# B&R Automation Studio project lab3
Automation Studio 4.5.2.102; technology packages: Acp10Arnc0 5.2.1

## Configuration Config1

CPU 4PP065.0571-P74, AutomationRuntime D4.52, Build 4.1.2, Vc V4.52.0, Safety 1.6

### Task classes (Cpu.sw)
```
Cyclic#1 (cycle 2000 us, tolerance 0 us):
  SDCAxisCtr <- SDCAxisCtrlX.prg
DataObjects: Acp10sys
NcDataObjects: acp10etxen <- acp10etxen.dob, Axis_Xa <- Axis_Xobj.Axis_Xa.dob, Axis_Xi <- Axis_Xobj.Axis_Xi.dob
Binaries: TCData, udbdef, ashwd, Role, User, sysconf, ashwac, asfw, arconfig, iomap, acp10cfg, Acp10map1, Acp10map
Libraries: Acp10man, Acp10par, NcGlobal, Acp10sdc, Acp10_MC, brsystem, sys_lib, runtime, AsBrStr, Acp10sim, AsIOTime, MotorContr, asstring, astime, fileio, powerlnk, asieccon
```

### Hardware
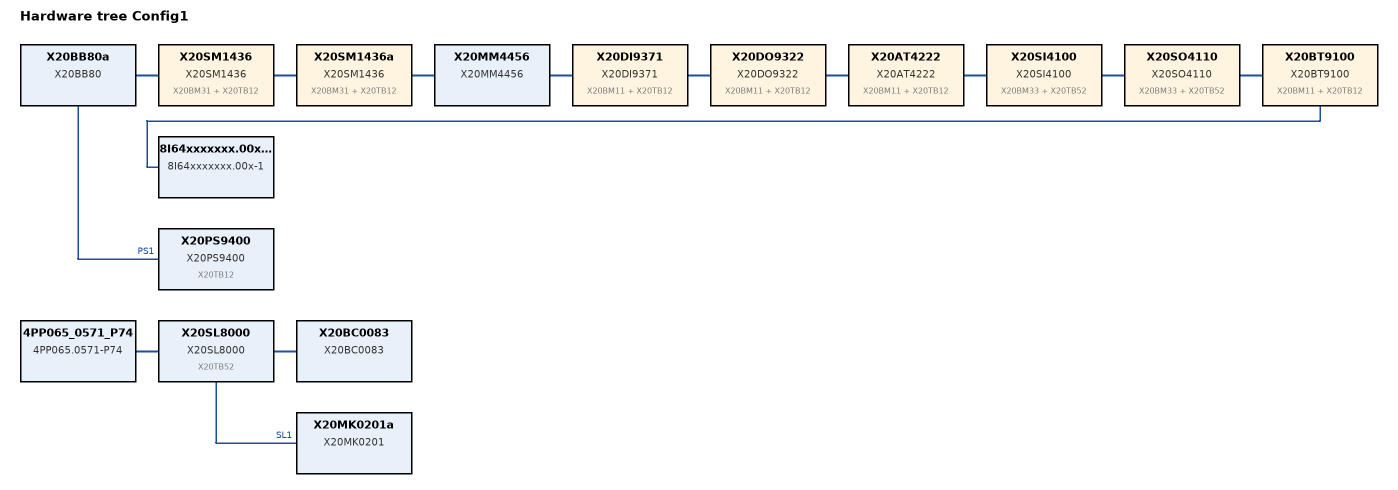
```
4PP065_0571_P74 : 4PP065.0571-P74 v1.1.2.0
  Connector IF5:
    ActivateDevice = 1
    Mode = Manual
    InternetAddress = 10.0.1.10
    SubnetMask = 255.255.255.0
  ConfigurationID = labBR
  TimerDeviceType = EPLX2X
  TimerDevice = 4PP065_0571_P74.IF4
  TaskClassIdleTime = 2000
  Cyclic1Duration = 2000
  Cyclic1Tolerance = 0
  Cyclic1Output = 1
8I64xxxxxxx.00x-1 : 8I64xxxxxxx.00x-1 v2.1.3.0  [X2X1 -> X20BT9100.X2X1 [Cable Type=X2XCable, Length=10, Version=1.0.0.2]]
  packedETAD = packed
  packedETI = packed
  packedCMDD = packed
  ACC = 30
  DEC = 30
  UNS = 220
  NCR = 10
  NSP = 890
  COS = 64
  RSC = 33000
X20AT4222 : X20AT4222 v1.2.3.0  [SS1 -> X20TB12f.SS; SL -> X20BM11c.SL1]
X20BB80a : X20BB80 v1.0.2.0
X20BC0083 : X20BC0083 v2.9.0.0  [PLK1 -> X20SL8000.PLK2 (NodeNumber=2) [Cable Type=PowerlinkCable, Length=10, Version=1.0.0.2]; SL -> X20BB80a.SL1]
X20BM11a : X20BM11 v1.0.0.1  [X2X1 -> X20MM4456.X2X2]
X20BM11b : X20BM11 v1.0.0.1  [X2X1 -> X20BM11a.X2X2]
X20BM11c : X20BM11 v1.0.0.1  [X2X1 -> X20BM11b.X2X2]
X20BM11d : X20BM11 v1.0.0.1  [X2X1 -> X20BM33b.X2X2]
X20BM31a : X20BM31 v1.0.0.1  [X2X1 -> X20BB80a.IF1]
X20BM31b : X20BM31 v1.0.0.1  [X2X1 -> X20BM31a.X2X2]
X20BM33a : X20BM33 v1.0.0.4  [X2X1 -> X20BM11c.X2X2]
X20BM33b : X20BM33 v1.0.0.4  [X2X1 -> X20BM33a.X2X2]
X20BT9100 : X20BT9100 v1.0.3.0  [SS1 -> X20TB12g.SS; SL -> X20BM11d.SL1]
X20DI9371 : X20DI9371 v1.0.2.0  [SS1 -> X20TB12d.SS; SL -> X20BM11a.SL1]
X20DO9322 : X20DO9322 v1.0.3.0  [SS1 -> X20TB12e.SS; SL -> X20BM11b.SL1]
X20MK0201a : X20MK0201 v1.0.0.0  [SL -> X20SL8000.SL1]
X20MM4456 : X20MM4456 v1.1.5.0  [X2X1 -> X20BM31b.X2X2]
X20PS9400 : X20PS9400 v1.8.0.0  [SS1 -> X20TB12b.SS; PS -> X20BB80a.PS1]
X20SI4100 : X20SI4100 v1.10.1.1  [SS1 -> X20TB52b.SS; SL -> X20BM33a.SL1]
X20SL8000 : X20SL8000 v1.6.5.2  [PLK1 -> 4PP065_0571_P74.IF4 (NodeNumber=1) [Cable Type=PowerlinkCable, Length=10, Version=1.0.0.2]; PLK2 -> X20BC0083.PLK1 (NodeNumber=1) [Cable Type=PowerlinkCable, Length=10, Version=1.0.0.2]; SS1 -> X20TB52a.SS]
  SafeProject = SafeLOGIC-1
  SafeDesigner = 3.0.18.3402403
X20SM1436 : X20SM1436 v2.3.0.0  [SS1 -> X20TB12a.SS; SL -> X20BM31a.SL1]
X20SM1436a : X20SM1436 v2.3.0.0  [SS1 -> X20TB12c.SS; SL -> X20BM31b.SL1]
X20SO4110 : X20SO4110 v1.10.1.1  [SS1 -> X20TB52c.SS; SL -> X20BM33b.SL1]
  SafeModuleID = 3
X20TB12a : X20TB12 v1.0.0.0
X20TB12b : X20TB12 v1.0.0.0
X20TB12c : X20TB12 v1.0.0.0
X20TB12d : X20TB12 v1.0.0.0
X20TB12e : X20TB12 v1.0.0.0
X20TB12f : X20TB12 v1.0.0.0
X20TB12g : X20TB12 v1.0.0.0
X20TB52a : X20TB52 v1.0.0.1
X20TB52b : X20TB52 v1.0.0.1
X20TB52c : X20TB52 v1.0.0.1
```

### IoMap.iom - 4PP065_0571_P74/IoMap.iom
```iecst
VAR_CONFIG
	::SDCAxisCtr:pwm_period AT %QW."X20MM4456".PeriodDurationPWM;
	::SDCAxisCtr:coil_pwm_value AT %QW."X20MM4456".PulseWidthCurrentPWM04;
	::SDCAxisCtr:pos_hand_btn AT %IX."X20DI9371".DigitalInput02;
	::SDCAxisCtr:neg_hand_btn AT %IX."X20DI9371".DigitalInput03;
	::SDCAxisCtr:coil_powered AT %IX."X20DI9371".DigitalInput01;
	::SDCAxisCtr:axis_X.pwm_value AT %QW."X20MM4456".PulseWidthCurrentPWM02;
	::SDCAxisCtr:axis_X.reset_error AT %QX."X20MM4456".ClearError02; (*Clear error motor bridge 01, clear endswitch*)
	::SDCAxisCtr:axis_X.reset_counter AT %QX."X20MM4456".ResetCounter02; (*Reset counter01 (1=reset active, 0=reset not active)*)
	::SDCAxisCtr:axis_X.endswitch_a_reached AT %IX."X20MM4456".StatusInput07; (*Logical condition input 03=Motor 01:R*)
	::SDCAxisCtr:axis_X.endswitch_b_reached AT %IX."X20MM4456".StatusInput08; (*Logical condition input 04=Motor 01:Reference enable/trigger/endswitch*)
	::SDCAxisCtr:axis_X.counter AT %IW."X20MM4456".Counter02; (*Count 01*)
END_VAR
```

### Acp10cfg.ncc - 4PP065_0571_P74/Motion/Acp10cfg.ncc
```
NcConfiguration (Version=5.02.1, NcSwId=Acp10)
  ACP10CF1_typ:
    cnt_nettrc_rec_drive = 1500
    bufsize_trace_upload = 1200
    tc_nc_man_task = Cyclic #1
    glob_pv_as_ncobject = Yes
    ncsys_dl_broadcast = Yes
    ncsys_dl_acp_reset = Yes
    safemc_log_err_to_ax = Yes
    network_init:
      ncsw_init_execute = Yes
      automatic_execute = No
      node_nr_warning = Yes
      net_err_before_ncact = Yes
    nettrc:
      enter_parsecrec = Yes
      enter_ncaction = Yes
      save_ring_startidx = Yes
    cam_prof_download:
      cam_dat_dl_parallel = No
      tc_cam_dl_parallel = Task class for NC Manager task
    sdc_if[0]:
      if_name = SDC_IF1
      mc_broadcast_size = 800
      mc_broadcast_extdat = No
```

### Acp10map1.ncm - 4PP065_0571_P74/Motion/Acp10map1.ncm
```
NcMapping (NcSwId=ACP10, DisabledNodesAreHidden=False)
  NcObject Axis_X (ModuleAddress=SDC_IF1.ST2, InterfaceType=SDC, Type=ncAXIS, Channel=1, AcoposSimulation=Off, InitParameter=Axis_Xi, AcoposParameter=Axis_Xa, Disabled=FALSE, ModuleDisabled=FALSE)
```

- Physical/Config1/4PP065_0571_P74/PvMap.vvm: same as Physical/Config1/4PP065_0571_P74/Cpu.per
## Logical view

Binary libraries used (declarations not repeated): operator, runtime, astime, AsIecCon, Acp10man 5.02.1, Acp10par 5.02.1, NcGlobal 5.02.1, Acp10sdc 5.02.1, Acp10_MC 5.02.1, brsystem, sys_lib, AsBrStr, Acp10sim 5.02.1, AsIOTime, asstring

### Global.var - Global variables
```iecst
VAR
	Axis_X : ACP10AXIS_typ;
	Axis_X_HW : SdcHwCfg_typ := (0);
	Axis_X_DrvIf : SdcDrvIf16_typ := (0);
	Axis_X_DiDoIf : SdcDiDoIf_typ := (0);
	Axis_X_ModuleOk : BOOL := 0;
	Axis_X_EncIf : SdcEncIf16_typ;
END_VAR
```

### Package Logical/Libraries - Global libraries

### Library Logical/Libraries/MotorContr (ANSIC)

#### MotorContr.fun - Exported functions and function blocks
```iecst
{REDUND_ERROR} {REDUND_UNREPLICABLE} FUNCTION_BLOCK FB_Integrator (*TODO: Add your comment here*) (*$GROUP=User,$CAT=User,$GROUPICON=User.png,$CATICON=User.png*)
	VAR_INPUT
		in : {REDUND_UNREPLICABLE} REAL;
	END_VAR
	VAR_OUTPUT
		out : {REDUND_UNREPLICABLE} REAL;
	END_VAR
	VAR
		dt : {REDUND_UNREPLICABLE} REAL;
	END_VAR
END_FUNCTION_BLOCK

{REDUND_ERROR} {REDUND_UNREPLICABLE} FUNCTION_BLOCK FB_Motor (*TODO: Add your comment here*) (*$GROUP=User,$CAT=User,$GROUPICON=User.png,$CATICON=User.png*)
	VAR_INPUT
		u : {REDUND_UNREPLICABLE} REAL; (*Напряжение на двигателе*)
	END_VAR
	VAR_OUTPUT
		w : {REDUND_UNREPLICABLE} REAL; (*Угловая скорость вала*)
		phi : {REDUND_UNREPLICABLE} REAL; (*Угол поворота вала*)
	END_VAR
	VAR
		integrator : {REDUND_UNREPLICABLE} FB_Integrator; (*Интегратор*)
		Tm : {REDUND_UNREPLICABLE} REAL; (*Механическая постоянная времени*)
		ke : {REDUND_UNREPLICABLE} REAL; (*коэф двигателя по напряжению*)
		dt : {REDUND_UNREPLICABLE} REAL; (*шаг дискретизации*)
	END_VAR
END_FUNCTION_BLOCK

{REDUND_ERROR} {REDUND_UNREPLICABLE} FUNCTION_BLOCK FB_Regulator (*TODO: Add your comment here*) (*$GROUP=User,$CAT=User,$GROUPICON=User.png,$CATICON=User.png*)
	VAR_INPUT
		e : {REDUND_UNREPLICABLE} REAL; (*ошибка регулирования*)
	END_VAR
	VAR_OUTPUT
		u : {REDUND_UNREPLICABLE} REAL; (*выходное напряжение*)
	END_VAR
	VAR
		k_p : {REDUND_UNREPLICABLE} REAL; (*кэф П-регулятора*)
		k_i : {REDUND_UNREPLICABLE} REAL; (*кэф И-регулятора*)
		integrator : {REDUND_UNREPLICABLE} FB_Integrator; (*интегратор*)
		iyOld : {REDUND_UNREPLICABLE} REAL; (*превышение выхода над ограничением*)
		max_abs_value : {REDUND_UNREPLICABLE} REAL; (*ограничение выхода*)
		dt : {REDUND_UNREPLICABLE} REAL; (*шаг дискретизации*)
	END_VAR
END_FUNCTION_BLOCK

{REDUND_ERROR} {REDUND_UNREPLICABLE} FUNCTION_BLOCK FB_Axis (*TODO: Add your comment here*) (*$GROUP=User,$CAT=User,$GROUPICON=User.png,$CATICON=User.png*)
	VAR_INPUT
		reset_error : {REDUND_UNREPLICABLE} BOOL; (*Сброс ошибок мотора*)
		endswitch_a_reached : {REDUND_UNREPLICABLE} BOOL; (*Состояние начального концевого датчика*)
		endswitch_b_reached : {REDUND_UNREPLICABLE} BOOL; (*Состояние конечного концевого датчика*)
	END_VAR
	VAR_OUTPUT
		reset_counter : {REDUND_UNREPLICABLE} BOOL; (*Сброс счётчика*)
		pwm_value : {REDUND_UNREPLICABLE} INT; (*Время Импулься ШИМ*)
		counter : {REDUND_UNREPLICABLE} INT; (*Счётчик импульсов*)
		speed : {REDUND_UNREPLICABLE} REAL; (*Скорость вращения оси двигателя*)
	END_VAR
	VAR
		last_counter : {REDUND_UNREPLICABLE} INT; (*Хранение предыдущего значения counter в процессе расчёта*)
		dt : {REDUND_UNREPLICABLE} REAL; (*Шаг дискретизации*)
	END_VAR
	VAR_INPUT
		u : {REDUND_UNREPLICABLE} REAL; (*Напряжение с выхода регулятора*)
	END_VAR
END_FUNCTION_BLOCK
```

#### FB_Integrator.c
```c
#include <bur/plctypes.h>
#ifdef __cplusplus
	extern "C"
	{
#endif
	#include "MotorContr.h"
#ifdef __cplusplus
	};
#endif
/* TODO: Add your comment here */
void FB_Integrator(struct FB_Integrator* inst)
{
	inst->out = inst->in * inst->dt + inst->out;
}
```

#### FB_Motor.c
```c
#include <bur/plctypes.h>
#ifdef __cplusplus
	extern "C"
	{
#endif
	#include "MotorContr.h"
#ifdef __cplusplus
	};
#endif
/* TODO: Add your comment here */
void FB_Motor(struct FB_Motor* inst)
{
	/*TODO: Add your code here*/
	inst->w = (inst->u / inst->ke - inst->w) * (inst->dt / inst->Tm) + inst->w;
	inst->integrator.in = inst->w * 3.1415f / 30.0f; // С переводом в [рад/с]
	inst->integrator.dt = inst->dt;
	FB_Integrator(&inst->integrator);
	inst->phi = inst->integrator.out;
}
```

#### FB_Regulator.c
```c
#include <bur/plctypes.h>
#ifdef __cplusplus
	extern "C"
	{
#endif
	#include "MotorContr.h"
#ifdef __cplusplus
	};
#endif
/* TODO: Add your comment here */
void FB_Regulator(struct FB_Regulator* inst)
{
	/*TODO: Add your code here*/
	float proportial = inst->e * inst->k_p;
	if (proportial > inst->max_abs_value)
	{
		proportial = inst->max_abs_value;
	}
	else if ( proportial < -inst->max_abs_value)
	{
		proportial = -inst->max_abs_value;
	}
	float integral_part_in = inst->e * inst->k_i - inst->iyOld / inst->dt;
	inst->integrator.in = integral_part_in;
	inst->integrator.dt = inst->dt;
	FB_Integrator(&inst->integrator);
	float sum = proportial + inst->integrator.out;

	if (sum > inst->max_abs_value)
	{
		inst->u = inst->max_abs_value;
	}
	else if (sum < -inst->max_abs_value)
	{
		inst->u = -inst->max_abs_value;
	}
	else inst->u = sum;

	inst->iyOld = sum - inst->u;
}
```

#### FB_Axis.c
```c
#include <bur/plctypes.h>
#ifdef __cplusplus
	extern "C"
	{
#endif
	#include "MotorContr.h"
#ifdef __cplusplus
	};
#endif
/* TODO: Add your comment here */
void FB_Axis(struct FB_Axis* inst)
{
	inst->pwm_value = (INT)(inst->u / 24.0f * 32767.0f);
	inst->speed = inst->u / 24.0f * 6500.0f;
}
```

### Data object Logical/acp10etxen (Ett)

- acp10etxen.ett (not shown)

### Package Logical/Axis_Xobj - Axis_Xobj

### Data object Logical/Axis_Xobj/Axis_Xa (Apt)

#### Axis_Xa.apt - Параметры инициализации оси
```
AcoposParameterTable:
  Root Parameters:
    109 = 24 (Name=SCALE_ENCOD_INCR)  // Encoder1: Encoder scaling: increments per encoder revolution
    64201 = 6500 (Name=SERVO_V_MAX_OUTPUT)
```

### Data object Logical/Axis_Xobj/Axis_Xi (Ax)

#### Axis_Xi.ax - Файл параметров инициализации оси
```
InitParameter (Version=5.02.1, NcSwId=ACP10)
  ACP10AXIS_typ:
    dig_in:
      level:
        reference = ncACTIV_HI
        pos_hw_end = ncACTIV_HI
        neg_hw_end = ncACTIV_HI
        trigger1 = ncACTIV_HI
        trigger2 = ncACTIV_HI
    encoder_if:
      parameter:
        count_dir = ncSTANDARD
        scaling:
          load:
            units = 3000
            rev_motor = 1
    limit:
      parameter:
        v_pos = 10000.0
        v_neg = 10000.0
        a1_pos = 10000.0
        a2_pos = 10000.0
        a1_neg = 10000.0
        a2_neg = 10000.0
        t_jolt = 0.0
        t_in_pos = 0.0
        pos_sw_end = 8388607
        neg_sw_end = -8388608
        ds_warning = 500.0
        ds_stop = 3000.0
        a_stop = 1.0E+30
        dv_stop = 0.0
        dv_stop_mode = ncOFF
    controller:
      mode = ncPOSITION
      position:
        kv = 10.0
        tn = 0.0
        t_predict = 0.01
        t_total = 0.01
        p_max = 1.0E+30
        i_max = 0.0
      speed:
        kv = 2.0
        tn = 0.0
        t_filter = 0.0
        isq_filter1:
          type = ncOFF
          a0 = 0.0
          a1 = 0.0
          b0 = 0.0
          b1 = 0.0
          b2 = 0.0
          c0_par_id = 0
          c1_par_id = 0
        isq_filter2:
          type = ncOFF
          a0 = 0.0
          a1 = 0.0
          b0 = 0.0
          b1 = 0.0
          b2 = 0.0
          c0_par_id = 0
          c1_par_id = 0
        isq_filter3:
          type = ncOFF
          a0 = 0.0
          a1 = 0.0
          b0 = 0.0
          b1 = 0.0
          b2 = 0.0
          c0_par_id = 0
          c1_par_id = 0
      uf:
        type = ncLINEAR + ncCORRECTION
        auto_config = ncMOTOR_PAR
        u0 = 0.0
        un = 0.0
        fn = 50.0
        k_f_slip = 0.0
      ff:
        torque_load = 0.0
        torque_pos = 0.0
        torque_neg = 0.0
        kv_torque = 0.0
        inertia = 0.0
        t_filter_a = 0.0
    move:
      stop:
        parameter[0]:
          decel_ramp = ncA_LIMIT
          controller = ncON
        parameter[1]:
          decel_ramp = ncA_LIMIT
          controller = ncON
        parameter[2]:
          decel_ramp = ncA_LIMIT
          controller = ncON
        parameter[3]:
          decel_ramp = ncA_LIMIT
          controller = ncON
        quickstop:
          decel_ramp = ncA_LIMIT
          t_jolt = 0.0
        drive_error:
          decel_ramp = ncA_LIMIT
      homing:
        parameter:
          s = 0
          v_switch = 2000.0
          v_trigger = 1600.0
          a = 10000.0
          mode = ncEND_SWITCH
          edge_sw = ncNEGATIVE
          start_dir = ncPOSITIVE
          trigg_dir = ncNEGATIVE
          ref_pulse = ncOFF
          fix_dir = ncOFF
          tr_s_block = 0.0
          torque_lim = 0.0
          ds_block = 0.0
          ds_stop = 0.0
      basis:
        parameter:
          v_pos = 2000.0
          v_neg = 2000.0
          a1_pos = 5000.0
          a2_pos = 5000.0
          a1_neg = 5000.0
          a2_neg = 5000.0
    message:
      text:
        parameter:
          format = ncBREAK
          columns = 80
          data_modul = acp10etxen
```

### Program Logical/SDCAxisCtrlX (ANSIC)

#### Main.c - Init, cyclic, exit code
```c
#include <bur/plctypes.h>

#ifdef _DEFAULT_INCLUDES
	#include <AsDefault.h>
#endif

void _INIT ProgramInit(void)
{
	axis_X.dt = 0.002f;

	Axis_X_HW.EncIf1_Typ = ncSDC_ENC16;
	Axis_X_HW.DiDoIf_Typ = ncSDC_DIDO;
	Axis_X_HW.DrvIf_Typ = ncSDC_DRVSERVO16;

	strcpy(Axis_X_HW.EncIf1_Name, "Axis_X_EncIf");
	strcpy(Axis_X_HW.DrvIf_Name, "Axis_X_DrvIf");
	strcpy(Axis_X_HW.DiDoIf_Name, "Axis_X_DiDoIf");
	Axis_X_EncIf.iEncOK = 1;
	Axis_X_DrvIf.iDrvOK = 1;
	Axis_X_DrvIf.iStatusEnable = 1;
	Axis_X_DiDoIf.iDriveReady = 1;

	fb_regulator.dt = 0.002f;
	//fb_motor.dt = 0.01f;
	//fb_motor.ke = 0.016f;
	//fb_motor.Tm = 0.1f;
	fb_regulator.max_abs_value = 24;
	fb_regulator.k_i = 0.16f;
	fb_regulator.k_p = 0.0f;
	fb_regulator.iyOld = 0.0f;

	axis_X.reset_error = 1;

	pwm_period = 200;
}

void _CYCLIC ProgramCyclic(void)
{
	BOOL ctrl_on;
	BOOL hand_pos;
	BOOL hand_neg;

	Axis_X_EncIf.iLifeCnt++;
	Axis_X_DiDoIf.iLifeCntDriveEnable++;
	Axis_X_DiDoIf.iLifeCntDriveReady++;
	Axis_X_DiDoIf.iLifeCntNegHwEnd++;
	Axis_X_DiDoIf.iLifeCntPosHwEnd++;
	Axis_X_DiDoIf.iLifeCntReference++;
	Axis_X_DrvIf.iLifeCnt++;
	Axis_X_EncIf.iActTime = (INT)AsIOTimeCyclicStart();

	Axis_X_EncIf.iActPos = axis_X.counter;
	Axis_X_DiDoIf.iPosHwEnd = axis_X.endswitch_a_reached;
	Axis_X_DiDoIf.iNegHwEnd = axis_X.endswitch_b_reached;
	Axis_X_DiDoIf.iDriveReady = coil_powered;

	coil_pwm_value = coil_powered ? 32767 : 0;

	ctrl_on = (Axis_X.controller.status == ncON);
	hand_pos = pos_hand_btn && !ctrl_on;
	hand_neg = neg_hand_btn && !ctrl_on;

	if (Axis_X.move.mode == ncHOMING)
		homing_active = 1;
	else if (homing_active && Axis_X.move.mode == ncOFF)
	{
		homing_active = 0;
		if (Axis_X.move.homing.status.ok && ctrl_on)
			ncaction((UDINT)&Axis_X, ncCONTROLLER, ncSWITCH_OFF);
	}

	fb_regulator.e = Axis_X_DrvIf.oSetPos * 6500.0f / 32767.0f - axis_X.speed;
	FB_Regulator(&fb_regulator);
	axis_X.u = fb_regulator.u;

	if (!coil_powered)
		axis_X.u = 0.0f;
	else if (hand_pos && !axis_X.endswitch_a_reached)
		axis_X.u = 12.0f;
	else if (hand_neg && !axis_X.endswitch_b_reached)
		axis_X.u = -12.0f;
	FB_Axis(&axis_X);
	if(axis_X.u > -4.0f && axis_X.u < 4.0f) // Слишком маленькое напряжение не позволяет провернуть двигатель, но пищит
		axis_X.pwm_value = 0;

	if (hand_pos || hand_neg || !coil_powered){
		axis_X.speed = 0.0f;
		fb_regulator.integrator.out = 0.0f;
		fb_regulator.iyOld = 0.0f;
	}
}

void _EXIT ProgramExit(void)
{

}
```

#### Variables.var - Local variables
```iecst
VAR
	homing_active : BOOL;
	axis_X : FB_Axis; (*Переменная оси*)
	coil_powered : BOOL; (*Включение обмотки возбуждения*)
	coil_pwm_value : INT; (*Время импулься ШИМ*)
	fb_motor : FB_Motor;
	fb_regulator : FB_Regulator; (*Переменная регулятора*)
	pwm_period : UINT; (*Период ШИМ*)
	fb_integrator : FB_Integrator;
	neg_hand_btn : BOOL;
	pos_hand_btn : BOOL;
END_VAR
```
